Fanuc KAREL source: ko00041.KL

-- PROVISIONAL review KL for V1013-1; original PC SHA256 ffb6ffa016045b3627ddf3c05683da785b9d0266f6922a9c7dd549e38c51202d
-- Incomplete behavior may be omitted. Consult companion uncertainty JSON. Do not deploy.
PROGRAM KO00041
%NOLOCKGROUP
BEGIN
  -- UNRESOLVED_PC offsets 5-12; opcodes 9D,23
  -- UNRESOLVED_PC offsets 17-69; opcodes 27,27,49,7E,AD,27,49,7E,AD,22,31,7E,4A
  -- UNRESOLVED_PC offsets 74-78; opcodes 7F
END KO00041
